SUBAPPLICATION Softkey_IXA_TO_logiBUS_QXA_BG (* Konvertierung Softkey IXA zu logiBUS QXA und Background *)
  (* Standard: 61499-2; Description: Copyright (c) 2023 Meisterschulen am Ostbahnhof This program and the accompanying materials are made available under the terms of the Eclipse Public License 2.0 which is available at https://www.eclipse.org/legal/epl-2.0/ SPDX-License-Identifier: EPL-2.0 *)
  (* Version 1.1, 2026-07-20, Franz Höpfinger, Meisterschulen am Ostbahnhof, Background *)
  (* Version 1.0, 2026-01-15, Franz Höpfinger, Meisterschulen am Ostbahnhof, initial API and implementation and/or initial documentation *)
  PACKAGE MyLib::sys;
  IMPORT isobus::UT::Q::const::IDs::ID_NULL;
  IMPORT logiBUS::io::DQ::logiBUS_DO;
  IMPORT logiBUS::io::DQ::logiBUS_DO_S;
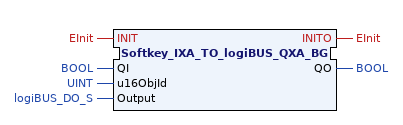
  EVENT_INPUT
    INIT : EInit; (* Initialization Request *)
  END_EVENT
  EVENT_OUTPUT
    INITO : EInit; (* Initialization Confirm *)
  END_EVENT
  VAR_INPUT
    QI : BOOL := TRUE; (* Quality Input - TRUE to enable service *)
    u16ObjId : UINT := ID_NULL; (* Object ID *)
    Output : logiBUS::io::DQ::logiBUS_DO_S := logiBUS_DO::Invalid; (* Identify the Output Output_Q1..Q8 *)
  END_VAR
  VAR_OUTPUT
    QO : BOOL; (* Quality Output - TRUE if service executed successfully *)
  END_VAR
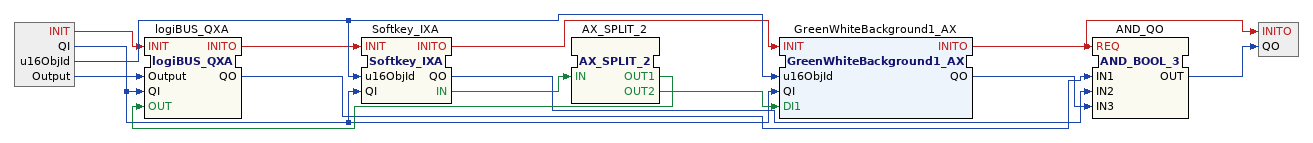
  FBS
    logiBUS_QXA : logiBUS::io::DQ::logiBUS_QXA;
    Softkey_IXA : isobus::UT::io::Softkey::Softkey_IXA;
    AX_SPLIT_2 : adapter::events::unidirectional::AX_SPLIT_2;
    AND_QO : iec61131::booleanOperators::AND_BOOL_3;
  END_FBS
  SUBAPPS
    GreenWhiteBackground1_AX : MyLib::sys::GreenWhiteBackground1_AX;
  END_SUBAPPS
  EVENT_CONNECTIONS
    INIT TO logiBUS_QXA.INIT;
    logiBUS_QXA.INITO TO Softkey_IXA.INIT;
    Softkey_IXA.INITO TO GreenWhiteBackground1_AX.INIT;
    GreenWhiteBackground1_AX.INITO TO INITO;
    GreenWhiteBackground1_AX.INITO TO AND_QO.REQ;
  END_CONNECTIONS
  DATA_CONNECTIONS
    u16ObjId TO Softkey_IXA.u16ObjId;
    Output TO logiBUS_QXA.Output;
    u16ObjId TO GreenWhiteBackground1_AX.u16ObjId;
    QI TO logiBUS_QXA.QI;
    QI TO Softkey_IXA.QI;
    logiBUS_QXA.QO TO AND_QO.IN1;
    Softkey_IXA.QO TO AND_QO.IN2;
    AND_QO.OUT TO QO;
    QI TO GreenWhiteBackground1_AX.QI;
    GreenWhiteBackground1_AX.QO TO AND_QO.IN3;
  END_CONNECTIONS
  ADAPTER_CONNECTIONS
    Softkey_IXA.IN TO AX_SPLIT_2.IN;
    AX_SPLIT_2.OUT1 TO logiBUS_QXA.OUT;
    AX_SPLIT_2.OUT2 TO GreenWhiteBackground1_AX.DI1;
  END_CONNECTIONS
END_SUBAPPLICATION
